(****************************************************************************************************<br>
© Syntegon Group.<br>
All rights reserved, also regarding any disposal, exploitation, reproduction, editing, distribution,<br>
as well as in the event of applications for industrial property rights.<br>
*****************************************************************************************************<br>
DESCRIPTION:<br>
Runs the TcUnit unit tests of the libraries Syn_Visu and Syn_Config (the installed SynVisu and SynConfig, newest<br>
versions) once after the start: every suite in POUs/Tests (_FB_TestConfig... for Syn_Config). TcUnit writes the<br>
results to the error list (ADS log) and, through TcUnit-Runner, to an xUnit file. Tests use only the libraries'<br>
public methods and their contract structures, written as the gateway writes them.<br>
****************************************************************************************************)
PROGRAM P_TestRun
VAR
	fb_TestComponent					: _FB_TestComponent;
	fb_TestConveyor						: _FB_TestConveyor;
	fb_TestProductRegister				: _FB_TestProductRegister;
	fb_TestRobot						: _FB_TestRobot;
	fb_TestXtsTrack						: _FB_TestXtsTrack;
	fb_TestBodyComponent				: _FB_TestBodyComponent;
	fb_TestMachine						: _FB_TestMachine;
	fb_TestConfigComponent				: _FB_TestConfigComponent;
	fb_TestConfigStaging				: _FB_TestConfigStaging;
	fb_TestConfigRobot					: _FB_TestConfigRobot;
	fb_TestConfigBodyComponent			: _FB_TestConfigBodyComponent;
	fb_TestConfigMachine				: _FB_TestConfigMachine;
	fb_TestConfigTopology				: _FB_TestConfigTopology;
END_VAR

TcUnit.RUN();

END_PROGRAM

(* stored: Version 1.1.0.1
   POU P_TestRun: Id {c2d649ca-bc8a-434d-92a6-238352d2fa0a}, SpecialFunc None *)
